(* IEC 61131-3 sources: ironplc/compiler/syntax/tests/fixtures/codesys, 11 files *)

(* ---- oop_members.st ---- *)
INTERFACE IStartable EXTENDS IRunnable, IStoppable
END_INTERFACE

FUNCTION_BLOCK ABSTRACT Motor EXTENDS Drive IMPLEMENTS IStartable, IStoppable
VAR_INPUT
    enable : BOOL;
END_VAR
VAR_OUTPUT
    running : BOOL;
END_VAR
VAR
    speed : REAL := 0.0;
END_VAR
running := enable;

METHOD PUBLIC FINAL Start : BOOL
VAR_INPUT
    target : REAL;
END_VAR
VAR_INST
    starts : INT;
END_VAR
starts := starts + 1;
speed := target;
Start := TRUE;
END_METHOD

METHOD ABSTRACT Stop
END_METHOD

PROPERTY Rpm : REAL
GET
    Rpm := speed * 60.0;
END_GET
SET
    speed := Rpm / 60.0;
END_SET
END_PROPERTY
END_FUNCTION_BLOCK

(* ---- sfc_chart.st ---- *)
FUNCTION_BLOCK Sequence
VAR_INPUT go : BOOL; END_VAR
INITIAL_STEP Idle:
    Light(N);
END_STEP
STEP Running:
    Light(N, lit);
    Pulse(SD, T#2s);
END_STEP
TRANSITION Start (PRIORITY := 1) FROM Idle TO Running := go; END_TRANSITION
TRANSITION FROM Running TO Idle := NOT go; END_TRANSITION
ACTION Light:
    lit := TRUE;
END_ACTION
END_FUNCTION_BLOCK

(* ---- configuration.st ---- *)
CONFIGURATION Plant
    VAR_GLOBAL
        shared : INT;
    END_VAR
    RESOURCE Cpu ON PLC
        VAR_GLOBAL
            local : BOOL;
        END_VAR
        TASK Fast (INTERVAL := T#10ms, PRIORITY := 1);
        TASK Slow (SINGLE := trigger, PRIORITY := 5);
        PROGRAM Main WITH Fast : Control (setpoint := 10, out => shared, Motor WITH Slow);
        PROGRAM RETAIN Aux : Logger;
    END_RESOURCE
    VAR_CONFIG
        Cpu.Main.motor.speed AT %QW0 : INT := 5;
    END_VAR
END_CONFIGURATION

(* ---- control_flow.st ---- *)
(* Loop control, jumps and the conditional statements of CODESYS, a direct
   address read in a statement, and a qualified enumeration value in the
   initial value of a structure. *)
TYPE
    Color : (Red, Green, Blue);
    Pair : STRUCT
        a : INT;
        b : Color;
    END_STRUCT;
    First : Pair := (a := 1, b := Color#Red);
END_TYPE

PROGRAM control_flow
VAR
    i : INT;
    total : INT;
    ready : BOOL;
    sensor : BOOL;
END_VAR
    sensor := %IX0.1;
    FOR i := 0 TO 10 DO
        IF i = 3 THEN
            CONTINUE;
        END_IF;
        IF i = 8 THEN
            EXIT;
        END_IF;
        total := total + i;
    END_FOR;
    WHILE ready DO
        EXIT;
    END_WHILE;
    JMP (ready) skip;
    total := 0;
skip:
    CALC (ready, notify(1));
    __WAIT(ready);
END_PROGRAM

(* ---- direct_variables.st ---- *)
PROGRAM IoDemo
VAR
    input_bit AT %IX0.0 : BOOL;
    output_word AT %QW1 : WORD;
    counter : DINT;
END_VAR
output_word := 16#00FF;
input_bit := FALSE;
END_PROGRAM

(* ---- namespaces.st ---- *)
NAMESPACE Outer
    TYPE Level : INT; END_TYPE
    NAMESPACE Inner
        FUNCTION Twice : INT
        VAR_INPUT x : INT; END_VAR
        Twice := x * 2;
        END_FUNCTION
    END_NAMESPACE
END_NAMESPACE

PROGRAM Main
END_PROGRAM

(* ---- pragmas.st ---- *)
{attribute 'strict'}
PROGRAM PragmaDemo
VAR
    counter : DINT;
END_VAR
counter := counter + 1;
END_PROGRAM

(* ---- references_and_pointers.st ---- *)
PROGRAM ReferenceDemo
VAR
    target : INT;
    alias : REFERENCE TO INT;
    raw_ptr : POINTER TO INT;
END_VAR
alias := target;
raw_ptr := ADR(target);
raw_ptr^ := target + 1;
END_PROGRAM

(* ---- strings_and_comments.st ---- *)
PROGRAM StringsDemo
VAR
    name : STRING(80);
    wide : WSTRING(40);
END_VAR
// a CODESYS-style line comment
name := 'Wärmebild';
(* a block comment *)
wide := "wide";
END_PROGRAM

(* ---- time_literals.st ---- *)
PROGRAM TimeDemo
VAR
    delay : TIME := T#1m30s;
    stamp : LTIME := LTIME#2h15m;
    timeout : TIME := T#250ms;
END_VAR
delay := delay + T#1s;
END_PROGRAM

(* ---- types_and_variables.st ---- *)
TYPE
    Percent : INT(0..100) := 50;
    Name : STRING[32] := 'pump';
    Wide : WSTRING(16);
    Vector : ARRAY[1..3] OF REAL := [1.0, 2.0, 3.0];
    Table : ARRAY[0..1, 0..2] OF INT;
    Open : ARRAY[*] OF BYTE;
    Color : (Red, Green := 5, Blue) BYTE := Green;
    Point : STRUCT
        x : INT := 1;
        y : INT := 2;
        label : STRING[8];
    END_STRUCT;
    Overlay : UNION
        whole : WORD;
        bytes : ARRAY[0..1] OF BYTE;
    END_UNION;
    Pen : Point := (x := 3, y := 4);
    IntRef : REF_TO INT;
    Alias : REFERENCE TO INT;
    Handle : POINTER TO DINT;
    Args : PARAMS(4) OF INT;
END_TYPE

VAR_GLOBAL CONSTANT
    Limit : INT := 10;
END_VAR

VAR_GLOBAL RETAIN
    counter : DINT;
    flag : BOOL;
END_VAR

PROGRAM Variables
VAR_INPUT
    start : BOOL R_EDGE;
    stop : BOOL F_EDGE;
END_VAR
VAR_IN_OUT
    shared : INT;
END_VAR
VAR RETAIN
    total : DINT := 0;
    zero, one : INT := 1;
END_VAR
VAR
    in_bit AT %IX0.0 : BOOL;
    words : ARRAY[1..4] OF INT := [4(0)];
    pen : Point := (x := 1, y := 2);
    motor : Fb(enable := TRUE);
    ptr : POINTER TO INT;
    target_ref : REF_TO INT := REF(total);
END_VAR
VAR_EXTERNAL CONSTANT
    Limit : INT;
END_VAR
VAR_STAT
    calls : INT;
END_VAR
total := total + 1;
END_PROGRAM
